(* IEC 61131-3 sources: lasal-git-demo/CPU/LasalDemoProject/Class/SdiasBase (part 2) *)

  elsif TempRetCode = ERROR then
    ret_code := ERROR;
  else
    ret_code := BUSY;
  end_if;

END_FUNCTION

FUNCTION VIRTUAL GLOBAL SdiasBase::GetDeviceID
	VAR_OUTPUT
		output 	: UDINT;
	END_VAR

  //Overwrite in derived Classes
  output := HWC_INVALID_DEVICE_ID;

END_FUNCTION

FUNCTION VIRTUAL SdiasBase::GetFWVersion
	VAR_INPUT
		pData 	: ^CHAR;
		Length 	: UDINT;
	END_VAR

  //Overwrite in derived Classes
  if pData then
    if Length >= 1 then
      pData^ := 0;    // Set first byte  to 0 termination = invalid string
    end_if;
  end_if;

END_FUNCTION

FUNCTION VIRTUAL GLOBAL SdiasBase::GetHWTimeStamp
	VAR_OUTPUT
		HWTimeStamp 	: UINT;
	END_VAR
  VAR
    MyPara   : CmdStruct;
    MyResult : results;
    retval   : iprStates;
  END_VAR

  HWTimeStamp := 0;

  MyPara.uiCmd := CMD_GET_HW_TIMESTAMP;
  MyPara.aPara[0]$t_GetHwTimestampCmd.udVersion    := 1;
  MyPara.aPara[0]$t_GetHwTimestampCmd.udCoreSelect := 0;

  retval := SdiasIn.NewInst(#MyPara, #MyResult);
  if retval = READY then
    if MyResult.uiLng >= sizeof(t_GetHwTimestampResult) then
      HWTimeStamp := MyResult.aData[0]$t_GetHwTimestampResult.uiTimeStamp;
    end_if;
  end_if;

END_FUNCTION

FUNCTION VIRTUAL GLOBAL SdiasBase::UpdateRtPreOp
#pragma warning(disable:0073);
	VAR_INPUT
		callinfo 	: t_SDIAS_UpdateRTPreOp;
	END_VAR
#pragma warning(default:0073);
	VAR_OUTPUT
		ret_code 	: iprStates;
	END_VAR

  // Overerload in derived Classes
//  case callinfo of
//  	t_SDIAS_UpdateRTPreOp::SDIAS_RTPREOP_CHECKSYNC:
//  	t_SDIAS_UpdateRTPreOp::SDIAS_RTPREOP_CHECKDATAVALID:
//  end_case;

  ret_code := READY;

END_FUNCTION
FUNCTION SdiasBase::AddDynRdAccess
	VAR_INPUT
		hOffset 	: HINT;
		uLength 	: UINT;
		bCtrlAcc0 	: BOOL;(* := false *)
		ppData 	: pVoid;
		ppStateByte 	: pVoid;
		ppControlByte 	: pVoid;
		pAccessHandle 	: ^UDINT;
		WaitForAccessHandle 	: UDINT;
	END_VAR
	VAR_OUTPUT
		ret_code 	: iprStates;
	END_VAR
  VAR
  	MyPara   : CmdStruct;
    MyResult : results;
  END_VAR

  MyPara.uiCmd := SDIAS_CMD_ADD_DYN_RD_ACCESS;
  MyPara.aPara[0] := this$DINT;
  MyPara.aPara[1] := Place$DINT;
  MyPara.aPara[2] := Required;
  MyPara.aPara[3] := hOffset;
  MyPara.aPara[4] := uLength;
  MyPara.aPara[5] := ppData$DINT;
  MyPara.aPara[6] := ppStateByte$DINT;
  MyPara.aPara[7] := ppControlByte$DINT;
  MyPara.aPara[8] := pAccessHandle$DINT;
  MyPara.aPara[9] := WaitForAccessHandle$DINT;
  MyPara.aPara[10]:= to_dint(bCtrlAcc0);

  ret_code := SdiasIn.NewInst(#MyPara, #MyResult);

  if ret_code <> READY then
    LogValue("@02C9 (SdiasBase::AddDynRdAccess) Failed to add read access for SDIAS module at Place 0x{0}, offset {1}", Place, to_udint(hOffset));
  end_if;

END_FUNCTION

FUNCTION SdiasBase::AddDynWrAccess
	VAR_INPUT
		hOffset 	: HINT;
		uLength 	: UINT;
		bCtrlAcc0 	: BOOL;(* := false *)
		ppData 	: pVoid;
		ppStateByte 	: pVoid;
		ppControlByte 	: pVoid;
		pAccessHandle 	: ^UDINT;
		WaitForAccessHandle 	: UDINT;
	END_VAR
	VAR_OUTPUT
		ret_code 	: iprStates;
	END_VAR
  VAR
  	MyPara   : CmdStruct;
    MyResult : results;
  END_VAR

  MyPara.uiCmd := SDIAS_CMD_ADD_DYN_WR_ACCESS;
  MyPara.aPara[0] := this$DINT;
  MyPara.aPara[1] := Place$DINT;
  MyPara.aPara[2] := Required;
  MyPara.aPara[3] := hOffset;
  MyPara.aPara[4] := uLength;
  MyPara.aPara[5] := ppData$DINT;
  MyPara.aPara[6] := ppStateByte$DINT;
  MyPara.aPara[7] := ppControlByte$DINT;
  MyPara.aPara[8] := pAccessHandle$DINT;
  MyPara.aPara[9] := WaitForAccessHandle$DINT;
  MyPara.aPara[10]:= to_dint(bCtrlAcc0);

  ret_code := SdiasIn.NewInst(#MyPara, #MyResult);

  if ret_code <> READY then
    LogValue("@02CA (SdiasBase::AddDynWrAccess) Failed to add write access for SDIAS module at Place 0x{0}, offset {1}", Place, to_udint(hOffset));
  end_if;

END_FUNCTION

FUNCTION SdiasBase::ChangeDynAccess
	VAR_INPUT
		AccessHandle 	: UDINT;
		NewOffset 	: HDINT;
		NewLength 	: UDINT;
	END_VAR
 	VAR_OUTPUT
		ret_code 	: iprStates;
	END_VAR
  VAR
  	MyPara   : CmdStruct;
    MyResult : results;
  END_VAR

  MyPara.uiCmd := SDIAS_CMD_CHANGE_DYN_ACCESS;
  MyPara.aPara[0] := AccessHandle$DINT;
  MyPara.aPara[1] := NewOffset$DINT;
  MyPara.aPara[2] := NewLength$DINT;
  ret_code := SdiasIn.NewInst(#MyPara, #MyResult);

  if ret_code <> READY then
    LogValue("@03F6 (SdiasBase::ChangeDynAccess) Failed to change access for SDIAS module at Place 0x{0}", Place);
  end_if;

END_FUNCTION

FUNCTION VIRTUAL SdiasBase::SPIWriteAddAccesses
	VAR_OUTPUT
		eModuleInitState 	: iprStates;
	END_VAR

  //This method has to be called in the derivated class if the class wants to use this feature

  //Add dynamic write access for write SPI Data
  if AddDynWrAccess(hOffset             := SDIAS_SPI_MASTER_ADRESS_TRANSMIT_BUFFER0
                 , uLength              := sizeof(t_SPI_PDO_DataWrite)
                 , bCtrlAcc0            := 1                                //Control Write Access
                 , ppData               := #sSPIVars.pWriteData
                 , ppStateByte          := #sSPIVars.sWriteAccess.pStateByte
                 , ppControlByte        := #sSPIVars.sWriteAccess.pControlByte
                 , pAccessHandle        := #sSPIVars.sWriteAccess.udAccessHandle
                 , WaitForAccessHandle  := 0
                 ) <> READY then

    LogError(pMsg:="@02ED (SdiasBase::SPIWriteAddAccesses) Adding dynamic write access for SPI Write functionality failed!");
    eModuleInitState := ERROR;
    return;
  end_if;

  //Add dynamic read access for reading SPI Data
  if AddDynRdAccess(hOffset             := SDIAS_SPI_MASTER_ADRESS_RECEIVE_BUFFER0
                 , uLength              := sizeof(t_SPI_PDO_DataRead)
                 , bCtrlAcc0            := 1                                //Control Read Access
                 , ppData               := #sSPIVars.pReadData
                 , ppStateByte          := #sSPIVars.sReadAccess.pStateByte
                 , ppControlByte        := #sSPIVars.sReadAccess.pControlByte
                 , pAccessHandle        := #sSPIVars.sReadAccess.udAccessHandle
                 , WaitForAccessHandle  := 0
                 ) <> READY then

    LogError(pMsg:="@02EE (SdiasBase::SPIWriteAddAccesses) Adding dynamic read access for SPI Write functionality failed!");
    eModuleInitState := ERROR;
    return;
  end_if;

  //Add dynamic read access for reading status of SPI Master
  if AddRdAccess(hOffset              := SDIAS_SPI_MASTER_ADRESS_STATUS_REGISTER
               , uLength              := 1
               , bCtrlAcc0            := 1                                //Control Read Access
               , ppData               := #sSPIVars.pReadStateData
               , ppStateByte          := #sSPIVars.sReadStateAccess.pStateByte
               , ppControlByte        := #sSPIVars.sReadStateAccess.pControlByte
               , pAccessHandle        := #sSPIVars.sReadStateAccess.udAccessHandle
               , WaitForAccessHandle  := 0
               ) <> READY then

    LogError(pMsg:="@02EE (SdiasBase::SPIWriteAddAccesses) Adding dynamic read access for SPI Write functionality failed!");
    eModuleInitState := ERROR;
    return;
  end_if;

  //if access are ok
  eModuleInitState := READY;

END_FUNCTION

FUNCTION VIRTUAL SdiasBase::SPIWriteGetState
	VAR_OUTPUT
		retcode	: iprStates;
	END_VAR

  //initialize return code with busy
  retcode := BUSY;

  if sSPIVars.bsFinished.Error then
    //error occured while write spi data
    retcode := ERROR;
  elsif sSPIVars.bsFinished.Finished then
    //write spi has finished
    retcode := READY;
  end_if;

END_FUNCTION

FUNCTION VIRTUAL SdiasBase::WriteSPIData
	VAR_INPUT
		usSectorNumber 	: USINT;
		usPageNumber 	: USINT;
		usPageOffset 	: USINT;
		udLength 	: UDINT;
		pData 	: ^USINT;
		usWriteMode 	: usWriteModes;(* := 0x00 *)
	END_VAR
	VAR_OUTPUT
		retcode 	: DINT;
	END_VAR

  retcode := 0;

  //Check for valid data
  if pData = nil then
    retcode := -1;
    return;
  end_if;

  //Check if last access finished or it was finished with error
  if sSPIVars.eSPIWriteSSW <> _SPIWrite_Idle then
    retcode := -2;
    return;
  end_if;

  //Check for valid length
  if udLength = 0 then
    retcode := -3;
    return;
  end_if;

  //Check if user write data is within the sector size
  if (((usPageNumber * SDIAS_SPI_PAGE_SIZE) + usPageOffset + udLength) > SDIAS_SPI_SECTOR_SIZE) then
    retcode := -4;
    return;
  end_if;

  //only access spi if it is locked
  if sSPIAccess.eSPIAccessProtect = _NotLocked then
    retcode := -5;
    return;
  end_if;

  sSPIVars.udUserWriteLength  := udLength;
  sSPIVars.usUserSectorNumber := usSectorNumber;
  sSPIVars.usUserPageNumber   := usPageNumber;
  sSPIVars.usUserPageOffset   := usPageOffset;
  sSPIVars.pUserWriteData     := pData;
  sSPIVars.usWriteMode        := usWriteMode;

  //reset error ssw
  sSPIVars.eSPIWriteSSWError := t_e_SPIWriteSSW::_SPIWrite_Idle;
  sSPIVars.bsFinished        := 0;

  case sSPIVars.usWriteMode of
    0,2:
      //read/write full sector
      sSPIVars.udMemoryToAllocate          := SDIAS_SPI_SECTOR_SIZE;
      sSPIVars.sReadAccess.usAccessLength  := SDIAS_MAX_PDO_SIZE;
      sSPIVars.sWriteAccess.usAccessLength := SDIAS_MAX_PDO_SIZE;
      sSPIVars.uiCurrentPage               := 0;
      sSPIVars.uiLastPage                  := SDIAS_SPI_PAGE_SIZE;
      sSPIVars.udUserDataOffset            := (sSPIVars.usUserPageNumber * SDIAS_SPI_PAGE_SIZE) + sSPIVars.usUserPageOffset;
    1,3:
      //read/write only required pages
      sSPIVars.udMemoryToAllocate          := ((sSPIVars.udUserWriteLength+SDIAS_SPI_PAGE_SIZE)/SDIAS_SPI_PAGE_SIZE)*SDIAS_SPI_PAGE_SIZE;
      sSPIVars.sReadAccess.usAccessLength  := SDIAS_MAX_PDO_SIZE/4;
      sSPIVars.sWriteAccess.usAccessLength := SDIAS_MAX_PDO_SIZE/4;
      sSPIVars.uiCurrentPage               := sSPIVars.usUserPageNumber;
      sSPIVars.uiLastPage                  := sSPIVars.uiCurrentPage + (sSPIVars.udUserWriteLength/SDIAS_SPI_PAGE_SIZE)$UINT + 1;
      sSPIVars.udUserDataOffset            := sSPIVars.usUserPageOffset;
  else
    retcode := -6;
    return;
  end_case;

  //allocate memory at SPIWriteUpdateCy()
  sSPIVars.eSPIWriteSSW   := t_e_SPIWriteSSW::_AllocateMemory;

END_FUNCTION

FUNCTION VIRTUAL SdiasBase::SPIWriteUpdateRt

  case sSPIVars.eSPIWriteSSW of

//*****************************************************************************
    t_e_SPIWriteSSW::_SPIWrite_Idle:
      //Wait for start
      //SSW will be set in method SPIWriteStart

//**********************************************************************************************************************************************************
//**********************************************************************************************************************************************************
//START REQUEST
//**********************************************************************************************************************************************************
//**********************************************************************************************************************************************************
  	t_e_SPIWriteSSW::_SetRequest:

      //Start/Stop data objects (is needed for the next steps)
      if sSPIVars.sWriteAccess.pControlByte then
        sSPIVars.sWriteAccess.pControlByte^.EnableDO := TRUE;
      else
        //error at start dataobject for spi access
        sSPIVars.eSPIWriteSSWError := sSPIVars.eSPIWriteSSW;
        sSPIVars.eSPIWriteSSW      := t_e_SPIWriteSSW::_ClearRequest;
        return;
      end_if;

      if sSPIVars.sReadAccess.pControlByte then
        sSPIVars.sReadAccess.pControlByte^.EnableDO := TRUE;
      else
        //error at start dataobject for spi access
        sSPIVars.eSPIWriteSSWError := sSPIVars.eSPIWriteSSW;
        sSPIVars.eSPIWriteSSW      := t_e_SPIWriteSSW::_ClearRequest;
        return;
      end_if;

      if sSPIVars.sReadStateAccess.pControlByte then
        sSPIVars.sReadStateAccess.pControlByte^.EnableDO := TRUE;
      else
        //error at start dataobject for spi access
        sSPIVars.eSPIWriteSSWError := sSPIVars.eSPIWriteSSW;
        sSPIVars.eSPIWriteSSW      := t_e_SPIWriteSSW::_ClearRequest;
        return;
      end_if;

      //Change write DO length
      ChangeDynAccess(AccessHandle :=  sSPIVars.sWriteAccess.udAccessHandle
                   , NewOffset    :=  SDIAS_SPI_MASTER_ADRESS_REQUEST_REGISTER
                   , NewLength    :=  1
                   );

      //Set Software request for SPI Master
      sSPIVars.pWriteData^[0] := SDIAS_SPI_MASTER_SOFTWARE_REQUEST;

      //Set length and offset for read object
      ChangeDynAccess(AccessHandle :=  sSPIVars.sReadAccess.udAccessHandle
                   , NewOffset    :=  SDIAS_SPI_MASTER_ADRESS_GRANT_REGISTER
                   , NewLength    :=  1
                   );

      sSPIVars.udTimeout    := ops.tAbsolute;
      sSPIVars.eSPIWriteSSW := t_e_SPIWriteSSW::_ReadGrant;

//*****************************************************************************
  	t_e_SPIWriteSSW::_ReadGrant:

      //Stop write object (is not needed for the next steps, will be enabled again if needed)
      sSPIVars.sWriteAccess.pControlByte^.EnableDO  := FALSE;

      //Check for grant
      if sSPIVars.pReadData^[0] = SDIAS_SPI_MASTER_SOFTWARE_REQUEST then

        //We got a grant, carry on
        //check if read of sector - page is needed
        case sSPIVars.usWriteMode of
          0,1:
            sSPIVars.eSPIWriteSSW := t_e_SPIWriteSSW::_ReadSectorData_SetPageAddress;
          2,3:
            //read of sector / page is not needed -> erase sector
            sSPIVars.eSPIWriteSSW := t_e_SPIWriteSSW::_EraseSector_SetPageAddress;
        end_case;
        sSPIVars.eSPIWriteSSW := t_e_SPIWriteSSW::_ReadSectorData_SetPageAddress;
      elsif (ops.tAbsolute-sSPIVars.udTimeout) >= SDIAS_SPI_TIMEOUT then
        //error at getting grant for spi access
        sSPIVars.eSPIWriteSSWError := sSPIVars.eSPIWriteSSW;
        sSPIVars.eSPIWriteSSW      := t_e_SPIWriteSSW::_ClearRequest;
      end_if;

//**********************************************************************************************************************************************************
//**********************************************************************************************************************************************************
//READ SECTOR DATA
//**********************************************************************************************************************************************************
//**********************************************************************************************************************************************************
  	t_e_SPIWriteSSW::_ReadSectorData_SetPageAddress:

      //Start write object (is needed for the next steps)
      sSPIVars.sWriteAccess.pControlByte^.EnableDO  := TRUE;

      ChangeDynAccess(AccessHandle :=  sSPIVars.sWriteAccess.udAccessHandle
                   , NewOffset    :=  SDIAS_SPI_MASTER_ADRESS_PAGE_ADRESS
                   , NewLength    :=  2
                   );

      //Due to the reason that we have to read the whole sector, just use the sector number from the user write address
      sSPIVars.pWriteData^[0]$UINT := (sSPIVars.usUserSectorNumber SHL 8) + sSPIVars.uiCurrentPage; //Byte 1 .. Pagenumber, Byte 2 .. Sectornumber

      sSPIVars.udTimeout    := ops.tAbsolute;
      sSPIVars.eSPIWriteSSW := t_e_SPIWriteSSW::_ReadSectorData_Wait4SetPageAddress;

//*****************************************************************************
  	t_e_SPIWriteSSW::_ReadSectorData_Wait4SetPageAddress:

      //Stop write object (is not needed for the next steps, will be enabled again if needed)
      sSPIVars.sWriteAccess.pControlByte^.EnableDO  := FALSE;

      if sSPIVars.pReadStateData^$USINT = SDIAS_SPI_MASTER_STATE_READY  then
        sSPIVars.eSPIWriteSSW := t_e_SPIWriteSSW::_ReadSectorData_SetReadPageCommand;
      elsif (ops.tAbsolute-sSPIVars.udTimeout) >= SDIAS_SPI_TIMEOUT then
        //timeout while waiting for spi master state ready
        sSPIVars.eSPIWriteSSWError := sSPIVars.eSPIWriteSSW;
        sSPIVars.eSPIWriteSSW      := t_e_SPIWriteSSW::_ClearRequest;
      end_if;

//*****************************************************************************
	  t_e_SPIWriteSSW::_ReadSectorData_SetReadPageCommand:

      //Start write object (is needed for the next steps)
      sSPIVars.sWriteAccess.pControlByte^.EnableDO  := TRUE;

      ChangeDynAccess(AccessHandle :=  sSPIVars.sWriteAccess.udAccessHandle
                   , NewOffset    :=  SDIAS_SPI_MASTER_ADRESS_PREDEFINED_COMMAND_REGISTER
                   , NewLength    :=  1
                   );

      sSPIVars.sReadAccess.usAccessOffset   := 0;
      sSPIVars.sWriteAccess.usAccessOffset  := 0;

      sSPIVars.pWriteData^$USINT := SDIAS_SPI_MASTER_COMMAND_PAGE_READ;

      ChangeDynAccess(AccessHandle :=  sSPIVars.sReadAccess.udAccessHandle
                   , NewOffset    :=  SDIAS_SPI_MASTER_ADRESS_RECEIVE_BUFFER0
                   , NewLength    :=  sSPIVars.sReadAccess.usAccessLength
                   );
      sSPIVars.udTimeout    := ops.tAbsolute;
      sSPIVars.eSPIWriteSSW := t_e_SPIWriteSSW::_ReadSectorData_Wait4SetReadPageCommand;

//*****************************************************************************
  	t_e_SPIWriteSSW::_ReadSectorData_Wait4SetReadPageCommand:

      //Stop write object (is not needed for the next steps, will be enabled again if needed)
      sSPIVars.sWriteAccess.pControlByte^.EnableDO  := FALSE;
      if sSPIVars.pReadStateData^$USINT = SDIAS_SPI_MASTER_STATE_READY  then
        sSPIVars.usCycleWaitCnt := 1;
        sSPIVars.eSPIWriteSSW   := t_e_SPIWriteSSW::_ReadSectorData_ReadReceiveBufferPart1;
      elsif (ops.tAbsolute-sSPIVars.udTimeout) >= SDIAS_SPI_TIMEOUT then
        //timeout while waiting for spi master state ready
        sSPIVars.eSPIWriteSSWError := sSPIVars.eSPIWriteSSW;
        sSPIVars.eSPIWriteSSW      := t_e_SPIWriteSSW::_ClearRequest;
      end_if;

//*****************************************************************************
  	t_e_SPIWriteSSW::_ReadSectorData_ReadReceiveBufferPart1:

      //Check if the module is connected via VARAN (behind a VI02x), so we have to wait an additional cycle until we can access the data
      if bIsConnectedViaVARAN then
        //ChangeDynAccess was done in last cycle, so in this cycle the access will be changed and in the next cycle we can access the data
        if sSPIVars.usCycleWaitCnt = 0 then
          sSPIVars.usCycleWaitCnt += 1;
          return;
        end_if;
        sSPIVars.usCycleWaitCnt := 0;
      end_if;

      //Read the first part of the receive buffer
      //Receive buffer is 256 byte huge but our read DO can only read maximal 128 Byte with one access -> split it into more accesses

      //Part 1: Copy Byte 0 to 127 from receive buffer
      _memcpy(ptr1:=sSPIVars.pSectorMemoryRead + sSPIVars.udCurrentSectorMemoryOffset + sSPIVars.sReadAccess.usAccessOffset, ptr2:= sSPIVars.pReadData, cntr:=sSPIVars.sReadAccess.usAccessLength);
      //Also copy it to write buffer
      _memcpy(ptr1:=sSPIVars.pSectorMemoryWrite + sSPIVars.udCurrentSectorMemoryOffset + sSPIVars.sReadAccess.usAccessOffset, ptr2:= sSPIVars.pReadData, cntr:=sSPIVars.sReadAccess.usAccessLength);

      sSPIVars.sReadAccess.usAccessOffset += sSPIVars.sReadAccess.usAccessLength;

      if sSPIVars.sReadAccess.usAccessOffset < SDIAS_MAX_PDO_SIZE then

        ChangeDynAccess(AccessHandle :=  sSPIVars.sReadAccess.udAccessHandle
                     , NewOffset    :=  SDIAS_SPI_MASTER_ADRESS_RECEIVE_BUFFER0+sSPIVars.sReadAccess.usAccessOffset
                     , NewLength    :=  sSPIVars.sReadAccess.usAccessLength
                     );

      else
        //Increment offset to copy data
        sSPIVars.udCurrentSectorMemoryOffset += sizeof(t_SPI_PDO_DataRead);

        ChangeDynAccess(AccessHandle :=  sSPIVars.sReadAccess.udAccessHandle
                     , NewOffset    :=  SDIAS_SPI_MASTER_ADRESS_RECEIVE_BUFFER1
                     , NewLength    :=  sSPIVars.sReadAccess.usAccessLength
                     );

        sSPIVars.sReadAccess.usAccessOffset := 0;
        sSPIVars.eSPIWriteSSW := t_e_SPIWriteSSW::_ReadSectorData_ReadReceiveBufferPart2;
      end_if;

//*****************************************************************************
  	t_e_SPIWriteSSW::_ReadSectorData_ReadReceiveBufferPart2:

      //Check if the module is connected via VARAN (behind a VI02x), so we have to wait an additional cycle until we can access the data
      if bIsConnectedViaVARAN then
        //ChangeDynAccess was done in last cycle, so in this cycle the access will be changed and in the next cycle we can access the data
        if sSPIVars.usCycleWaitCnt = 0 then
          sSPIVars.usCycleWaitCnt += 1;
          return;
        end_if;
        sSPIVars.usCycleWaitCnt := 0;
      end_if;

      //Part 2: Copy Byte 128 to 255 from receive buffer
      _memcpy(ptr1:=sSPIVars.pSectorMemoryRead + sSPIVars.udCurrentSectorMemoryOffset+ sSPIVars.sReadAccess.usAccessOffset, ptr2:= sSPIVars.pReadData, cntr:=sSPIVars.sReadAccess.usAccessLength);

      //Also copy it to write buffer
      _memcpy(ptr1:=sSPIVars.pSectorMemoryWrite + sSPIVars.udCurrentSectorMemoryOffset + sSPIVars.sReadAccess.usAccessOffset, ptr2:= sSPIVars.pReadData, cntr:=sSPIVars.sReadAccess.usAccessLength);

      sSPIVars.sReadAccess.usAccessOffset += sSPIVars.sReadAccess.usAccessLength;

      if sSPIVars.sReadAccess.usAccessOffset < SDIAS_MAX_PDO_SIZE then

        ChangeDynAccess(AccessHandle :=  sSPIVars.sReadAccess.udAccessHandle
                     , NewOffset    :=  SDIAS_SPI_MASTER_ADRESS_RECEIVE_BUFFER1+sSPIVars.sReadAccess.usAccessOffset
                     , NewLength    :=  sSPIVars.sReadAccess.usAccessLength
                     );

      else
        //Increment offset to copy data
        sSPIVars.udCurrentSectorMemoryOffset += sizeof(t_SPI_PDO_DataRead);

        //Increment every page we read
        sSPIVars.uiCurrentPage               += 1;
        sSPIVars.sReadAccess.usAccessOffset  := 0;

        //Check if we have read the last page
        if sSPIVars.uiCurrentPage = sSPIVars.uiLastPage then

          sSPIVars.eSPIWriteSSW := t_e_SPIWriteSSW::_EraseSector_SetPageAddress;

          //Stop ReadDo (is not needed for the next steps, will be enabled again if needed)
          sSPIVars.sReadAccess.pControlByte^.EnableDO := FALSE;

        else
          sSPIVars.eSPIWriteSSW := t_e_SPIWriteSSW::_ReadSectorData_SetPageAddress;
        end_if;
      end_if;

//**********************************************************************************************************************************************************
//**********************************************************************************************************************************************************
//ERASE SECTOR
//**********************************************************************************************************************************************************
//**********************************************************************************************************************************************************
	t_e_SPIWriteSSW::_EraseSector_SetPageAddress:

      //Reset our page/sector counters
      case sSPIVars.usWriteMode of
        0,2:
          sSPIVars.uiCurrentPage := 0;
        1,3:
          sSPIVars.uiCurrentPage := sSPIVars.usUserPageNumber;
      end_case;
      sSPIVars.udCurrentSectorMemoryOffset := 0;

      //copy user data into memory write buffer
      _memcpy(ptr1 := sSPIVars.pSectorMemoryWrite + sSPIVars.udUserDataOffset
            , ptr2 := sSPIVars.pUserWriteData
            , cntr := sSPIVars.udUserWriteLength);

      //Start write object (is needed for the next steps)
      sSPIVars.sWriteAccess.pControlByte^.EnableDO  := TRUE;

      ChangeDynAccess(AccessHandle :=  sSPIVars.sWriteAccess.udAccessHandle
                   , NewOffset    :=  SDIAS_SPI_MASTER_ADRESS_PAGE_ADRESS
                   , NewLength    :=  2
                   );

      sSPIVars.udTimeout           := ops.tAbsolute;
      sSPIVars.pWriteData^[0]$UINT := (sSPIVars.usUserSectorNumber SHL 8);
      sSPIVars.eSPIWriteSSW        := t_e_SPIWriteSSW::_EraseSector_Wait4SetPageAddress;

//*****************************************************************************
	t_e_SPIWriteSSW::_EraseSector_Wait4SetPageAddress:

      //Stop write object (is not needed for the next steps, will be enabled again if needed)
      sSPIVars.sWriteAccess.pControlByte^.EnableDO  := FALSE;

      if sSPIVars.pReadStateData^$USINT = SDIAS_SPI_MASTER_STATE_READY  then
        sSPIVars.eSPIWriteSSW := t_e_SPIWriteSSW::_EraseSector_SetEraseSectorCommand;
      elsif (ops.tAbsolute-sSPIVars.udTimeout) >= SDIAS_SPI_TIMEOUT then
        //timeout while waiting for spi master state ready
        sSPIVars.eSPIWriteSSWError := sSPIVars.eSPIWriteSSW;
        sSPIVars.eSPIWriteSSW      := t_e_SPIWriteSSW::_ClearRequest;
      end_if;

//*****************************************************************************
  	t_e_SPIWriteSSW::_EraseSector_SetEraseSectorCommand:

      //Start write object (is needed for the next steps)
      sSPIVars.sWriteAccess.pControlByte^.EnableDO  := TRUE;

      ChangeDynAccess(AccessHandle :=  sSPIVars.sWriteAccess.udAccessHandle
                   , NewOffset    :=  SDIAS_SPI_MASTER_ADRESS_PREDEFINED_COMMAND_REGISTER
                   , NewLength    :=  1
                   );

      sSPIVars.udTimeout         := ops.tAbsolute;
      sSPIVars.pWriteData^$USINT := SDIAS_SPI_MASTER_COMMAND_SECTOR_ERASE;
      sSPIVars.eSPIWriteSSW      := t_e_SPIWriteSSW::_EraseSector_Wait4SetEraseSectorCommand;

//*****************************************************************************
  	t_e_SPIWriteSSW::_EraseSector_Wait4SetEraseSectorCommand:

      //Stop write object (is not needed for the next steps, will be enabled again if needed)
      sSPIVars.sWriteAccess.pControlByte^.EnableDO  := FALSE;

      if sSPIVars.pReadStateData^$USINT = SDIAS_SPI_MASTER_STATE_READY  then
        sSPIVars.eSPIWriteSSW := t_e_SPIWriteSSW::_WriteSectorData_SetPageAddress;
      elsif (ops.tAbsolute-sSPIVars.udTimeout) >= SDIAS_SPI_TIMEOUT then
        //timeout while waiting for spi master state ready
        sSPIVars.eSPIWriteSSWError := sSPIVars.eSPIWriteSSW;
        sSPIVars.eSPIWriteSSW      := t_e_SPIWriteSSW::_ClearRequest;
      end_if;

//**********************************************************************************************************************************************************
//**********************************************************************************************************************************************************
//WRITE SECTOR DATA
//**********************************************************************************************************************************************************
//**********************************************************************************************************************************************************
    t_e_SPIWriteSSW::_WriteSectorData_SetPageAddress:

      //Start write object (is needed for the next steps)
      sSPIVars.sWriteAccess.pControlByte^.EnableDO  := TRUE;

      //Wait until last write/erase sector has finished
      ChangeDynAccess(AccessHandle :=  sSPIVars.sWriteAccess.udAccessHandle
                   , NewOffset    :=  SDIAS_SPI_MASTER_ADRESS_PAGE_ADRESS
                   , NewLength    :=  2
                   );

      //Due to the reason that we have to write the whole sector, just use the sector number from the user write address
      sSPIVars.pWriteData^[0]$UINT := (sSPIVars.usUserSectorNumber SHL 8) + sSPIVars.uiCurrentPage;
      sSPIVars.udTimeout           := ops.tAbsolute;
      sSPIVars.eSPIWriteSSW        := t_e_SPIWriteSSW::_WriteSectorData_Wait4SetPageAddress;

//*****************************************************************************
    t_e_SPIWriteSSW::_WriteSectorData_Wait4SetPageAddress:

      //Stop write object (is not needed for the next steps, will be enabled again if needed)
      sSPIVars.sWriteAccess.pControlByte^.EnableDO  := FALSE;

      if sSPIVars.pReadStateData^$USINT = SDIAS_SPI_MASTER_STATE_READY  then
        sSPIVars.sWriteAccess.usAccessOffset := 0;
        sSPIVars.eSPIWriteSSW := t_e_SPIWriteSSW::_WriteSectorData_WriteTransmitBufferPart1;
      elsif (ops.tAbsolute-sSPIVars.udTimeout) >= SDIAS_SPI_TIMEOUT then
        //timeout while waiting for spi master state ready
        sSPIVars.eSPIWriteSSWError := sSPIVars.eSPIWriteSSW;
        sSPIVars.eSPIWriteSSW      := t_e_SPIWriteSSW::_ClearRequest;
      end_if;

//*****************************************************************************
    t_e_SPIWriteSSW::_WriteSectorData_WriteTransmitBufferPart1:

      //Start write object (is needed for the next steps)
      sSPIVars.sWriteAccess.pControlByte^.EnableDO  := TRUE;

      //Write whole sector to SPI Flash
      ChangeDynAccess(AccessHandle :=  sSPIVars.sWriteAccess.udAccessHandle
                   , NewOffset    :=  SDIAS_SPI_MASTER_ADRESS_TRANSMIT_BUFFER0 + sSPIVars.sWriteAccess.usAccessOffset
                   , NewLength    :=  sSPIVars.sWriteAccess.usAccessLength
                   );

      //Copy sector write memory to Dataobject data
      _memcpy(ptr1:= sSPIVars.pWriteData
            , ptr2:= sSPIVars.pSectorMemoryWrite + sSPIVars.udCurrentSectorMemoryOffset + sSPIVars.sWriteAccess.usAccessOffset
            , cntr:= sSPIVars.sWriteAccess.usAccessLength
            );

      sSPIVars.sWriteAccess.usAccessOffset += sSPIVars.sWriteAccess.usAccessLength;

      if sSPIVars.sWriteAccess.usAccessOffset >= SDIAS_MAX_PDO_SIZE then
        sSPIVars.sWriteAccess.usAccessOffset := 0;
        sSPIVars.eSPIWriteSSW := t_e_SPIWriteSSW::_WriteSectorData_WriteTransmitBufferPart2;
      end_if;

//*****************************************************************************
    t_e_SPIWriteSSW::_WriteSectorData_WriteTransmitBufferPart2:

      //Write whole sector to SPI Flash
      ChangeDynAccess(AccessHandle :=  sSPIVars.sWriteAccess.udAccessHandle
                   , NewOffset    :=  SDIAS_SPI_MASTER_ADRESS_TRANSMIT_BUFFER1 + sSPIVars.sWriteAccess.usAccessOffset
                   , NewLength    :=  sSPIVars.sWriteAccess.usAccessLength
                   );

      //Copy sector write memory to Dataobject data
      _memcpy(ptr1:= sSPIVars.pWriteData
            , ptr2:= sSPIVars.pSectorMemoryWrite + sSPIVars.udCurrentSectorMemoryOffset + SDIAS_MAX_PDO_SIZE + sSPIVars.sWriteAccess.usAccessOffset
            , cntr:= sSPIVars.sWriteAccess.usAccessLength
            );

      sSPIVars.sWriteAccess.usAccessOffset += sSPIVars.sWriteAccess.usAccessLength;

      if sSPIVars.sWriteAccess.usAccessOffset >= SDIAS_MAX_PDO_SIZE then
        sSPIVars.sWriteAccess.usAccessOffset := 0;
        sSPIVars.eSPIWriteSSW := t_e_SPIWriteSSW::_WriteSectorData_SetWritePageCommand;
      end_if;

//*****************************************************************************
    t_e_SPIWriteSSW::_WriteSectorData_SetWritePageCommand:

      ChangeDynAccess(AccessHandle :=  sSPIVars.sWriteAccess.udAccessHandle
                   , NewOffset    :=  SDIAS_SPI_MASTER_ADRESS_PREDEFINED_COMMAND_REGISTER
                   , NewLength    :=  1
                   );
      sSPIVars.pWriteData^$USINT := SDIAS_SPI_MASTER_COMMAND_PAGE_PROGRAM;

      sSPIVars.udTimeout    := ops.tAbsolute;
      sSPIVars.eSPIWriteSSW := t_e_SPIWriteSSW::_WriteSectorData_Wait4SetWritePageCommand;

//*****************************************************************************
    t_e_SPIWriteSSW::_WriteSectorData_Wait4SetWritePageCommand:

      //Stop write object (is not needed for the next steps, will be enabled again if needed)
      sSPIVars.sWriteAccess.pControlByte^.EnableDO  := FALSE;

      if sSPIVars.pReadStateData^$USINT = SDIAS_SPI_MASTER_STATE_READY then

        //Increment page counter if program was OK
        sSPIVars.uiCurrentPage += 1;
        //Increment our offset
        sSPIVars.udCurrentSectorMemoryOffset += SDIAS_SPI_PAGE_SIZE;
        //reset retry counter
        sSPIVars.usRetryCnt   := 0;

        //Check if finished
        if sSPIVars.uiCurrentPage = sSPIVars.uiLastPage then
          sSPIVars.eSPIWriteSSW := t_e_SPIWriteSSW::_VerifySectorData_SetPageAddress;

          //Reset our page/sector counters
          case sSPIVars.usWriteMode of
            0,2:
              sSPIVars.uiCurrentPage := 0;
            1,3:
              sSPIVars.uiCurrentPage := sSPIVars.usUserPageNumber;
          end_case;

          sSPIVars.udCurrentSectorMemoryOffset := 0;

        else
          sSPIVars.eSPIWriteSSW := t_e_SPIWriteSSW::_WriteSectorData_SetPageAddress;
        end_if;
      elsif (ops.tAbsolute-sSPIVars.udTimeout) >= SDIAS_SPI_TIMEOUT then
        //timeout while waiting for spi master state ready
        sSPIVars.eSPIWriteSSW := t_e_SPIWriteSSW::_WriteSectorData_SetPageAddress;
        sSPIVars.usRetryCnt   += 1;
        if sSPIVars.usRetryCnt > SDIAS_SPI_WRITE_MAX_RETRIES then
          //reset retry counter
          sSPIVars.usRetryCnt        := 0;
          //timeout while waiting for spi master state ready
          sSPIVars.eSPIWriteSSWError := sSPIVars.eSPIWriteSSW;
          sSPIVars.eSPIWriteSSW      := t_e_SPIWriteSSW::_ClearRequest;
        end_if;
        sSPIVars.NotReadyCnt += 1;
      end_if;

//**********************************************************************************************************************************************************
//**********************************************************************************************************************************************************
//VERIFY SECTOR DATA
//**********************************************************************************************************************************************************
//**********************************************************************************************************************************************************
    t_e_SPIWriteSSW::_VerifySectorData_SetPageAddress:

      //Start write object (is needed for the next steps)
      sSPIVars.sWriteAccess.pControlByte^.EnableDO  := TRUE;

      ChangeDynAccess(AccessHandle :=  sSPIVars.sWriteAccess.udAccessHandle
                   , NewOffset    :=  SDIAS_SPI_MASTER_ADRESS_PAGE_ADRESS
                   , NewLength    :=  2
                   );

      //Due to the reason that we have to read the whole sector, just use the sector number from the user write address
      sSPIVars.pWriteData^[0]$UINT := (sSPIVars.usUserSectorNumber SHL 8) + sSPIVars.uiCurrentPage;
      sSPIVars.udTimeout    := ops.tAbsolute;
      sSPIVars.eSPIWriteSSW := t_e_SPIWriteSSW::_VerifySectorData_Wait4SetPageAddress;

//*****************************************************************************
    t_e_SPIWriteSSW::_VerifySectorData_Wait4SetPageAddress:

      //Stop write object (is not needed for the next steps, will be enabled again if needed)
      sSPIVars.sWriteAccess.pControlByte^.EnableDO  := FALSE;

      if sSPIVars.pReadStateData^$USINT = SDIAS_SPI_MASTER_STATE_READY  then
        sSPIVars.eSPIWriteSSW := t_e_SPIWriteSSW::_VerifySectorData_SetReadPageCommand;
      elsif (ops.tAbsolute-sSPIVars.udTimeout) >= SDIAS_SPI_TIMEOUT then
        //error at getting grant for spi access
        sSPIVars.eSPIWriteSSWError := sSPIVars.eSPIWriteSSW;
        sSPIVars.eSPIWriteSSW      := t_e_SPIWriteSSW::_ClearRequest;
      end_if;

//*****************************************************************************
    t_e_SPIWriteSSW::_VerifySectorData_SetReadPageCommand:

      //Start write object (is needed for the next steps)
      sSPIVars.sWriteAccess.pControlByte^.EnableDO  := TRUE;

      ChangeDynAccess(AccessHandle :=  sSPIVars.sWriteAccess.udAccessHandle
                   , NewOffset    :=  SDIAS_SPI_MASTER_ADRESS_PREDEFINED_COMMAND_REGISTER
                   , NewLength    :=  1
                   );

      sSPIVars.pWriteData^$USINT := SDIAS_SPI_MASTER_COMMAND_PAGE_READ;

      //Start ReadDo (is needed for the next steps)
      sSPIVars.sReadAccess.pControlByte^.EnableDO := TRUE;

      ChangeDynAccess(AccessHandle :=  sSPIVars.sReadAccess.udAccessHandle
                   , NewOffset    :=  SDIAS_SPI_MASTER_ADRESS_RECEIVE_BUFFER0
                   , NewLength    :=  sSPIVars.sReadAccess.usAccessLength
                   );

      sSPIVars.udTimeout    := ops.tAbsolute;
      sSPIVars.eSPIWriteSSW := t_e_SPIWriteSSW::_VerifySectorData_Wait4SetReadPageCommand;

//*****************************************************************************
    t_e_SPIWriteSSW::_VerifySectorData_Wait4SetReadPageCommand:

      //Stop write object (is not needed for the next steps, will be enabled again if needed)
      sSPIVars.sWriteAccess.pControlByte^.EnableDO  := FALSE;

      if sSPIVars.pReadStateData^$USINT = SDIAS_SPI_MASTER_STATE_READY  then
        sSPIVars.sReadAccess.usAccessOffset := 0;
        sSPIVars.usCycleWaitCnt := 1;
        sSPIVars.eSPIWriteSSW   := t_e_SPIWriteSSW::_VerifySectorData_ReadReceiveBufferPart1;
      elsif (ops.tAbsolute-sSPIVars.udTimeout) >= SDIAS_SPI_TIMEOUT then
        //error at getting grant for spi access
        sSPIVars.eSPIWriteSSWError := sSPIVars.eSPIWriteSSW;
        sSPIVars.eSPIWriteSSW      := t_e_SPIWriteSSW::_ClearRequest;
      end_if;

//*****************************************************************************
  	t_e_SPIWriteSSW::_VerifySectorData_ReadReceiveBufferPart1:

      //Check if the module is connected via VARAN (behind a VI02x), so we have to wait an additional cycle until we can access the data
      if bIsConnectedViaVARAN then
        //ChangeDynAccess was done in last cycle, so in this cycle the access will be changed and in the next cycle we can access the data
        if sSPIVars.usCycleWaitCnt = 0 then
          sSPIVars.usCycleWaitCnt += 1;
          return;
        end_if;
        sSPIVars.usCycleWaitCnt := 0;
      end_if;

      //Read the first part of the receive buffer
      //Receive buffer is 256 byte huge but our read DO can only read 128 Byte with one access -> split it into two accesses

      //Part 1: Copy Byte 0 to 127 from receive buffer
      _memcpy(ptr1:=sSPIVars.pSectorMemoryVerify + sSPIVars.udCurrentSectorMemoryOffset + sSPIVars.sReadAccess.usAccessOffset, ptr2:= sSPIVars.pReadData, cntr:=sSPIVars.sReadAccess.usAccessLength);

      sSPIVars.sReadAccess.usAccessOffset += sSPIVars.sReadAccess.usAccessLength;

      if sSPIVars.sReadAccess.usAccessOffset < SDIAS_MAX_PDO_SIZE then

        ChangeDynAccess(AccessHandle :=  sSPIVars.sReadAccess.udAccessHandle
                     , NewOffset    :=  SDIAS_SPI_MASTER_ADRESS_RECEIVE_BUFFER0+sSPIVars.sReadAccess.usAccessOffset
                     , NewLength    :=  sSPIVars.sReadAccess.usAccessLength
                     );

      else
        //Increment offset to copy data
        sSPIVars.udCurrentSectorMemoryOffset += sizeof(t_SPI_PDO_DataRead);

        ChangeDynAccess(AccessHandle :=  sSPIVars.sReadAccess.udAccessHandle
                     , NewOffset    :=  SDIAS_SPI_MASTER_ADRESS_RECEIVE_BUFFER1
                     , NewLength    :=  sSPIVars.sReadAccess.usAccessLength
                     );
        sSPIVars.sReadAccess.usAccessOffset := 0;
        sSPIVars.usCycleWaitCnt := 0;
        sSPIVars.eSPIWriteSSW   := t_e_SPIWriteSSW::_VerifySectorData_ReadReceiveBufferPart2;
      end_if;

//*****************************************************************************
  	t_e_SPIWriteSSW::_VerifySectorData_ReadReceiveBufferPart2:

      //Check if the module is connected via VARAN (behind a VI02x), so we have to wait an additional cycle until we can access the data
      if bIsConnectedViaVARAN then
        //ChangeDynAccess was done in last cycle, so in this cycle the access will be changed and in the next cycle we can access the data
        if sSPIVars.usCycleWaitCnt = 0 then
          sSPIVars.usCycleWaitCnt += 1;
          return;
        end_if;
        sSPIVars.usCycleWaitCnt := 0;
      end_if;

      //Part 2: Copy Byte 128 to 255 from receive buffer
      _memcpy(ptr1:=sSPIVars.pSectorMemoryVerify + sSPIVars.udCurrentSectorMemoryOffset+ sSPIVars.sReadAccess.usAccessOffset, ptr2:= sSPIVars.pReadData, cntr:=sSPIVars.sReadAccess.usAccessLength);

      sSPIVars.sReadAccess.usAccessOffset += sSPIVars.sReadAccess.usAccessLength;

      if sSPIVars.sReadAccess.usAccessOffset < SDIAS_MAX_PDO_SIZE then

        ChangeDynAccess(AccessHandle :=  sSPIVars.sReadAccess.udAccessHandle
                     , NewOffset    :=  SDIAS_SPI_MASTER_ADRESS_RECEIVE_BUFFER1+sSPIVars.sReadAccess.usAccessOffset
                     , NewLength    :=  sSPIVars.sReadAccess.usAccessLength
                     );

      else
        //next step at SPIWriteUpdateCy()
        sSPIVars.eSPIWriteSSW := _VerifySectorData_CompareData;
      end_if;

//*****************************************************************************
    t_e_SPIWriteSSW::_VerifySectorData_CompareData:
    //at SPIWriteUpdateCy()

//**********************************************************************************************************************************************************
//FINISH SPI WRITE
//**********************************************************************************************************************************************************
  	t_e_SPIWriteSSW::_ClearRequest:

      //Start write object (is needed for the next steps)
      if sSPIVars.sWriteAccess.pControlByte then
        sSPIVars.sWriteAccess.pControlByte^.EnableDO := TRUE;
      else
        //error at start dataobject for spi access
        sSPIVars.eSPIWriteSSW      := t_e_SPIWriteSSW::_DisableDataObjects;
        return;
      end_if;

      //Change write DO length
      ChangeDynAccess(AccessHandle :=  sSPIVars.sWriteAccess.udAccessHandle
                   , NewOffset    :=  SDIAS_SPI_MASTER_ADRESS_CLEAR_REQUEST_REGISTER
                   , NewLength    :=  1
                   );

      //Clear Software request for SPI Master
      sSPIVars.pWriteData^[0] := SDIAS_SPI_MASTER_SOFTWARE_REQUEST;

      sSPIVars.eSPIWriteSSW := _DisableDataObjects;

//*****************************************************************************
  	t_e_SPIWriteSSW::_DisableDataObjects:
      //Disable Data objects because they are not used anymore (will be enabled with next start of SPI write access)
      if sSPIVars.sWriteAccess.pControlByte then
        sSPIVars.sWriteAccess.pControlByte^.EnableDO := FALSE;
      end_if;
      if sSPIVars.sReadAccess.pControlByte then
        sSPIVars.sReadAccess.pControlByte^.EnableDO := FALSE;
      end_if;
      if sSPIVars.sReadStateAccess.pControlByte then
        sSPIVars.sReadStateAccess.pControlByte^.EnableDO := FALSE;
      end_if;
      //free memory at SPIWriteUpdateCy()
      sSPIVars.eSPIWriteSSW := _FreeMemory;

//*****************************************************************************
  	t_e_SPIWriteSSW::_FinishSPIWrite:

      //Reset SSW
      sSPIVars.eSPIWriteSSW := _SPIWrite_Idle;
      //spi write has finished
      sSPIVars.bsFinished.Finished := 1;
      //check if an error occured while spi write
      if sSPIVars.eSPIWriteSSWError <> sSPIVars.eSPIWriteSSW then
        //error occurred while spi access - act error step is saved at sSPIVars.eSPIWriteSSWError
        sSPIVars.bsFinished.Error := 1;
      end_if;

//*****************************************************************************
  end_case;

END_FUNCTION

FUNCTION VIRTUAL SdiasBase::SPIWriteUpdateCy

  case sSPIVars.eSPIWriteSSW of
//*****************************************************************************
    t_e_SPIWriteSSW::_SPIWrite_Idle:
      //Wait for start
      //SSW will be set in method WriteSPIData()

//**********************************************************************************************************************************************************
  	t_e_SPIWriteSSW::_AllocateMemory:

      //check pointer, if it's not nil it must be freed
      if sSPIVars.pSectorMemoryRead then
        ToStdLib.Free(mptr:=sSPIVars.pSectorMemoryRead);
        sSPIVars.pSectorMemoryRead := NIL;
      end_if;
      //Allocate memory for read sector (1 sector has 64kByte)
      sSPIVars.pSectorMemoryRead$^void    := ToStdLib.Malloc(size:=sSPIVars.udMemoryToAllocate);
      if sSPIVars.pSectorMemoryRead = NIL then
        LogError(pMsg:="@02EF (SdiasBase::SPIWriteUpdateCy) Failed to allocate memory for sSPIVars.pSectorMemoryRead.");
        //error at allocate memory for spi access
        sSPIVars.eSPIWriteSSWError := sSPIVars.eSPIWriteSSW;
        //next step at SPIWriteUpdateRt()
        sSPIVars.eSPIWriteSSW      := t_e_SPIWriteSSW::_ClearRequest;
        return;
      end_if;

      //check pointer, if it's not nil it must be freed
      if sSPIVars.pSectorMemoryWrite then
        ToStdLib.Free(mptr:=sSPIVars.pSectorMemoryWrite);
        sSPIVars.pSectorMemoryWrite := NIL;
      end_if;
      //Allocate memory for write sector (1 sector has 64kByte)
      sSPIVars.pSectorMemoryWrite$^void   := ToStdLib.Malloc(size:=sSPIVars.udMemoryToAllocate);
      if sSPIVars.pSectorMemoryWrite = NIL then
        LogError(pMsg:="@02F0 (SdiasBase::SPIWriteUpdateCy) Failed to allocate memory for sSPIVars.pSectorMemoryWrite.");
        //error at allocate memory for spi access
        sSPIVars.eSPIWriteSSWError := sSPIVars.eSPIWriteSSW;
        //next step at SPIWriteUpdateRt()
        sSPIVars.eSPIWriteSSW      := t_e_SPIWriteSSW::_ClearRequest;
        return;
      end_if;

      //check pointer, if it's not nil it must be freed
      if sSPIVars.pSectorMemoryVerify then
        ToStdLib.Free(mptr:=sSPIVars.pSectorMemoryVerify);
        sSPIVars.pSectorMemoryVerify := NIL;
      end_if;
      //Allocate memory for verify sector (1 sector has 64kByte)
      sSPIVars.pSectorMemoryVerify$^void  := ToStdLib.Malloc(size:=sSPIVars.udMemoryToAllocate);

      if sSPIVars.pSectorMemoryVerify = NIL then
        LogError(pMsg:="@02F1 (SdiasBase::SPIWriteUpdateCy) Failed to allocate memory for sSPIVars.pSectorMemoryVerify.");
        //error at allocate memory for spi access
        sSPIVars.eSPIWriteSSWError := sSPIVars.eSPIWriteSSW;
        //next step at SPIWriteUpdateRt()
        sSPIVars.eSPIWriteSSW      := t_e_SPIWriteSSW::_ClearRequest;
        return;
      end_if;

      //Clear the memory
      _memset(sSPIVars.pSectorMemoryRead,   16#FF, sSPIVars.udMemoryToAllocate);
      _memset(sSPIVars.pSectorMemoryWrite,  16#FF, sSPIVars.udMemoryToAllocate);
      _memset(sSPIVars.pSectorMemoryVerify, 16#FF, sSPIVars.udMemoryToAllocate);

      //next step at SPIWriteUpdateRt()
      sSPIVars.eSPIWriteSSW := t_e_SPIWriteSSW::_SetRequest;

//**********************************************************************************************************************************************************
//other steps are at SPIWriteUpdateRt()
//**********************************************************************************************************************************************************

//*****************************************************************************
    t_e_SPIWriteSSW::_VerifySectorData_CompareData:

      //Check if data is the same
      if _memcmp(ptr1:= sSPIVars.pSectorMemoryVerify + sSPIVars.udCurrentSectorMemoryOffset - sizeof(t_SPI_PDO_DataRead),
                 ptr2:= sSPIVars.pSectorMemoryWrite + sSPIVars.udCurrentSectorMemoryOffset - sizeof(t_SPI_PDO_DataRead),
                 cntr:=SDIAS_SPI_PAGE_SIZE) <> 0 then

        //Error
        sSPIVars.usRetryCnt += 1;

        //Reset our page/sector counters
        case sSPIVars.usWriteMode of
          0,2:
            sSPIVars.uiCurrentPage := 0;
          1,3:
            sSPIVars.uiCurrentPage := sSPIVars.usUserPageNumber;
        end_case;
        sSPIVars.udCurrentSectorMemoryOffset := 0;

        if sSPIVars.usRetryCnt > SDIAS_SPI_WRITE_MAX_RETRIES then
          sSPIVars.usRetryCnt   :=  0;
          //next step at SPIWriteUpdateRt()
          sSPIVars.eSPIWriteSSW := _ClearRequest;
        else
          sSPIVars.bsFinished   := 0;
          //next step at SPIWriteUpdateRt()
          sSPIVars.eSPIWriteSSW := _ReadSectorData_SetPageAddress;
        end_if;
      else
        //Increment offset to copy data
        sSPIVars.udCurrentSectorMemoryOffset += sizeof(t_SPI_PDO_DataRead);

        //Increment every page we read
        sSPIVars.uiCurrentPage               += 1;

        //Check if we have read the last page
        if sSPIVars.uiCurrentPage = sSPIVars.uiLastPage then
          //Data is equal, finish SPI communication
          //next step at SPIWriteUpdateRt()
          sSPIVars.eSPIWriteSSW := t_e_SPIWriteSSW::_ClearRequest;
        else
          //next step at SPIWriteUpdateRt()
          sSPIVars.eSPIWriteSSW := t_e_SPIWriteSSW::_VerifySectorData_SetPageAddress;
        end_if;
      end_if;

//**********************************************************************************************************************************************************
  	t_e_SPIWriteSSW::_FreeMemory:
      //Free memory
      if sSPIVars.pSectorMemoryRead then
        ToStdLib.Free(mptr:=sSPIVars.pSectorMemoryRead);
        sSPIVars.pSectorMemoryRead := NIL;
      end_if;
      if sSPIVars.pSectorMemoryWrite then
        ToStdLib.Free(mptr:=sSPIVars.pSectorMemoryWrite);
        sSPIVars.pSectorMemoryWrite := NIL;
      end_if;
      if sSPIVars.pSectorMemoryVerify then
        ToStdLib.Free(mptr:=sSPIVars.pSectorMemoryVerify);
        sSPIVars.pSectorMemoryVerify := NIL;
      end_if;

      sSPIVars.uiCurrentPage                := 0;
      sSPIVars.udCurrentSectorMemoryOffset  := 0;
       //next step at SPIWriteUpdateRt()
      sSPIVars.eSPIWriteSSW := _FinishSPIWrite;

//**********************************************************************************************************************************************************
  	t_e_SPIWriteSSW::_FinishSPIWrite:
    //at SPIWriteUpdateRt()

  end_case;

END_FUNCTION

FUNCTION SdiasBase::LockSPIAccess
	VAR_INPUT
		udAccessID 	: UDINT;
	END_VAR
	VAR_OUTPUT
		dRetCode 	: iprStates;
	END_VAR
  VAR
  	udTempVar : UDINT;
  END_VAR

  udTempVar := sigclib_atomic_cmpxchgU32(pValue:=#sSPIAccess.eSPIAccessProtect$UDINT, cmpVal:=_NotLocked, newVal:=udAccessID);

  if (udTempVar = 0) | (udTempVar = udAccessID) then
    //access to spi interface is granted
    sSPIAccess.udSPILastLockTime := ops.tAbsolute;
    dRetCode := READY;
  else
    //spi access is locked by another instance
    dRetCode := BUSY;
    if (ops.tAbsolute-sSPIAccess.udSPILastLockTime) > (SDIAS_SPI_LOCK_TIMEOUT*udBusTime*SDIAS_MAX_PDO_SIZE/(1000*sSPIVars.sWriteAccess.usAccessLength)) then
      //reset all accesses
      sSPIAccess.eSPIAccessProtect := _NotLocked;
      //reset spi SSW
      eGetSPIDataSSW := _GetDataObjectList;
      eGetObjectListSSW := _GetObjList;
    end_if;
  end_if;

END_FUNCTION

FUNCTION SdiasBase::UnlockSPIAccess
  VAR_INPUT
    udAccessID 	: UDINT;
  END_VAR
  VAR_OUTPUT
    dRetCode 	: iprStates;
  END_VAR

  //reset lock bit if compare value is ok
  sigclib_atomic_cmpxchgU32(pValue:=#sSPIAccess.eSPIAccessProtect$UDINT, cmpVal:=udAccessID, newVal:=_NotLocked);
  dRetCode := READY;

END_FUNCTION
